// TIA Portal V15.1 export
FUNCTION "MCP_RC_R5FCM" : Void   // FC9834, LAD
{ S7_Optimized_Access := 'TRUE' }
   VAR_INPUT
      "a" : Bool;
      "b" : Int;
   END_VAR
BEGIN
END_FUNCTION
